RoboDK station: Car_Painting_Cell_v16.rdk

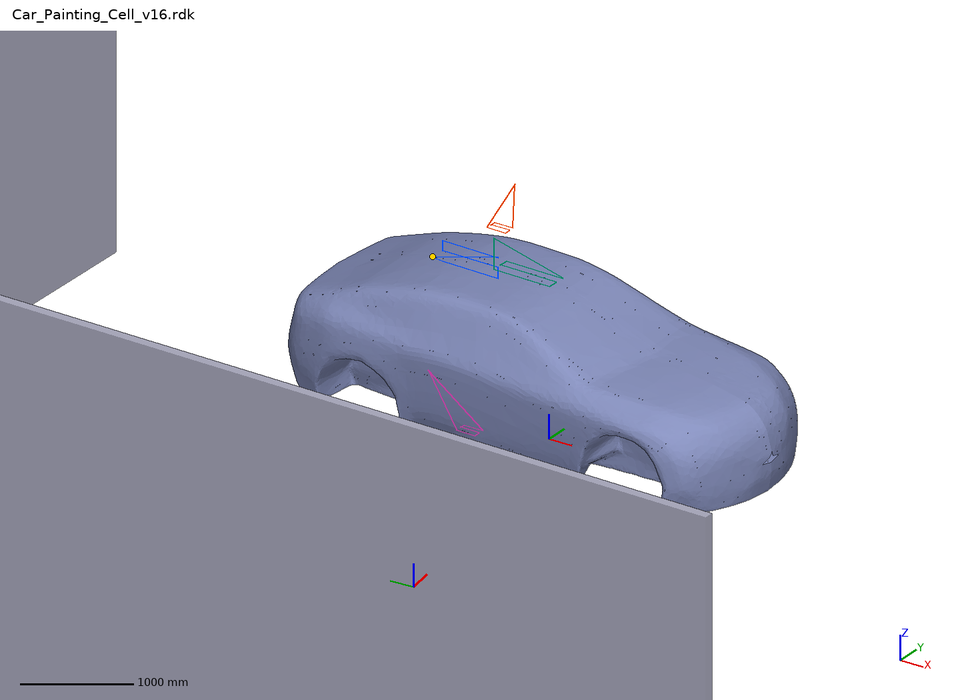
[picture v0: the station drawn from its stored meshes, robots at their saved joint values, targets as dots, program paths as lines]
Station Car_Painting_Cell_v16 (saved by RoboDK 6.1.1). Poses are relative to the parent item; angles as X-Y-Z fixed-axis rotations.
  - frame ABB IRB 6700-235/2.65 Base at (0, 0, 0) mm, rotated rx 1.67 ry -4.75 rz 96.19 deg
    - robot ABB IRB 6700-235/2.65: 6 axes, payload 235 kg, reach 2650 mm, repeatability 0.05 mm, weight 1280 kg
        joint limits [-170, -65, -180, -300, -130, -360] to [170, 85, 70, 300, 130, 360]; home [0, 0, 0, 0, 0, 0]; saved at [22.213, -18.762, 12.242, 0, 96.52, 202.213]
      - tool Generic Paint Sprayer, TCP at (50, 0, 450) mm, rotated rx 0 ry 30 rz 0 deg, size 277.6 x 203.2 x 501.7 mm
  - object Wall_Back at (0, -4050, 2000) mm, size 12000 x 100 x 4000 mm, geometry from Wall_Back.stl
  - object Wall_Side at (-6050, 0, 2000) mm, size 100 x 8000 x 4000 mm, geometry from Wall_Side.stl
  - frame Car_Frame at (-258.38, 2438.18, 404.41) mm
    - object Car_Body at (2438.35, -1259.55, -51.4) mm, rotated rx 0 ry 0 rz 90 deg, size 1981.5 x 4799.5 x 1349.6 mm, geometry from Sedan Car Body.IGS
  - Python program Setup_Cell (listed below)
  - program Paint_Side5 (10 instructions, listed below)
  - program Paint_Trunk2 (10 instructions, listed below)
  - program Paint_Roof2 (10 instructions, listed below)
  - program Paint_Hood2 (10 instructions, listed below)
  - program Main_Program (5 instructions, listed below)
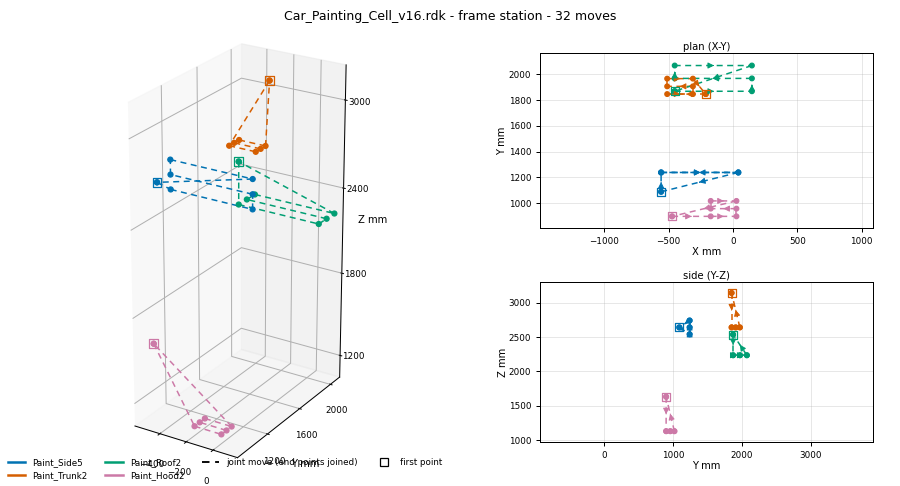
[picture p0: tool path of Car_Painting_Cell_v16.rdk in frame station, 32 of 35 moves have a stored position in this frame; points joined in program order, loops and branches not executed]

--- Python program Setup_Cell ---
# Type help("robodk.robolink") or help("robodk.robomath") for more information
# Press F5 to run the script
# Documentation: https://robodk.com/doc/en/RoboDK-API.html
# Reference:     https://robodk.com/doc/en/PythonAPI/robodk.html
# Note: It is not required to keep a copy of this file, your Python script is saved with your RDK project

# You can also use the new version of the API:
from robodk import robolink    # RoboDK API
from robodk import robomath    # Robot toolbox
RDK = robolink.Robolink()

# Forward and backwards compatible use of the RoboDK API:
# Remove these 2 lines to follow python programming guidelines
from robodk import *      # RoboDK API
from robolink import *    # Robot toolbox
# Link to RoboDK
# RDK = Robolink()

# Notify user:
print('To edit this program:\nright click on the Python program, then, select "Edit Python script"')

# Program example:
item = RDK.Item('base')
if item.Valid():
    print('Item selected: ' + item.Name())
    print('Item posistion: ' + repr(item.Pose()))

print('Items in the station:')
itemlist = RDK.ItemList()
print(itemlist)

# Provoking an exception will display the console output if you run this script from RoboDK
raise Exception('Program not edited.')

--- program Paint_Side5 (robot ABB IRB 6700-235/2.65) ---
  Set Ref.: Car_Frame
  Set Tool: Generic Paint Sprayer
  MoveJ 2 to (-300, -1350, 2235.34) mm, rotated rx -168.9 ry 64.7 rz -87.2 deg; joints [28.216, -32.938, 21.44, 101.638, -42.225, -113.719]
  MoveJ 3 to (-300, -1200, 2135.34) mm, rotated rx -168.9 ry 64.7 rz -87.2 deg; joints [23.122, -28.793, 24.985, 93.784, -36.162, -102.736]
  MoveJ 4 to (300, -1200, 2135.34) mm, rotated rx -168.9 ry 64.7 rz -87.2 deg; joints [-15.84, -33.97, 26.391, 23.272, 7.322, -30.496]
  MoveJ 5 to (300, -1200, 2235.34) mm, rotated rx -168.9 ry 64.7 rz -87.2 deg; joints [-15.495, -31.919, 20.419, 13.499, 10.949, -20.661]
  MoveJ 6 to (-300, -1200, 2235.34) mm, rotated rx -168.9 ry 64.7 rz -87.2 deg; joints [23.087, -26.983, 19.068, 99.337, -36.598, -109.625]
  MoveJ 7 to (-300, -1200, 2335.34) mm, rotated rx -168.9 ry 64.7 rz -87.2 deg; joints [23.052, -24.869, 12.83, 104.706, -37.424, -116.339]
  MoveJ 8 to (300, -1200, 2335.34) mm, rotated rx -168.9 ry 64.7 rz -87.2 deg; joints [-15.156, -29.592, 14.142, 8.67, 14.765, -15.792]
  MoveJ 9 to (-300, -1350, 2235.34) mm, rotated rx -168.9 ry 64.7 rz -87.2 deg; joints [28.216, -32.938, 21.44, 101.638, -42.225, -113.719]

--- program Paint_Trunk2 (robot ABB IRB 6700-235/2.65) ---
  Set Ref.: Car_Frame
  Set Tool: Generic Paint Sprayer
  MoveJ 2 to (47.14, -590.89, 2735.34) mm, rotated rx 176.1 ry 64.7 rz -87.2 deg; joints [-6.92, 10.197, -37.991, 14.59, 28.576, -12.875]
  MoveJ 3 to (-252.86, -590.89, 2235.34) mm, rotated rx 176.1 ry 64.7 rz -87.2 deg; joints [4.168, -2.249, 2.16, -88.78, 4.169, 88.777]
  MoveJ 4 to (-52.86, -590.89, 2235.34) mm, rotated rx 176.1 ry 64.7 rz -87.2 deg; joints [-3.705, -3.302, 2.796, 82.241, 3.739, -82.224]
  MoveJ 5 to (-52.86, -530.89, 2235.34) mm, rotated rx 176.1 ry 64.7 rz -87.2 deg; joints [-3.81, -0.342, 0.158, 87.229, 3.815, -87.223]
  MoveJ 6 to (-252.86, -530.89, 2235.34) mm, rotated rx 176.1 ry 64.7 rz -87.2 deg; joints [3.756, 0.675, -0.495, 87.264, -3.761, -87.258]
  MoveJ 7 to (-252.86, -470.89, 2235.34) mm, rotated rx 176.1 ry 64.7 rz -87.2 deg; joints [3.375, 3.631, -3.327, 84.87, -3.388, -84.861]
  MoveJ 8 to (-52.86, -470.89, 2235.34) mm, rotated rx 176.1 ry 64.7 rz -87.2 deg; joints [-3.908, 2.644, -2.656, 89.824, 3.908, -89.824]
  MoveJ 9 to (47.14, -590.89, 2735.34) mm, rotated rx 176.1 ry 64.7 rz -87.2 deg; joints [-6.92, 10.197, -37.991, 14.59, 28.576, -12.875]

--- program Paint_Roof2 (robot ABB IRB 6700-235/2.65) ---
  Set Ref.: Car_Frame
  Set Tool: Generic Paint Sprayer
  MoveJ 2 to (-194.48, -569.09, 2130.93) mm, rotated rx 176.1 ry 64.7 rz -87.2 deg; joints [12.275, 4.238, -19.199, -40.125, 19.263, 38.507]
  MoveJ 3 to (-194.48, -569.09, 1830.93) mm, rotated rx 176.1 ry 64.7 rz -87.2 deg; joints [12.149, -1.74, 1.882, 89.341, -12.15, -89.326]
  MoveJ 4 to (405.52, -569.09, 1830.93) mm, rotated rx 176.1 ry 64.7 rz -87.2 deg; joints [-11.823, -4.921, 3.782, 84.574, 11.877, -84.456]
  MoveJ 5 to (405.52, -469.09, 1830.93) mm, rotated rx 176.1 ry 64.7 rz -87.2 deg; joints [-11.459, -0.017, -0.535, 87.282, 11.472, -87.227]
  MoveJ 6 to (-194.48, -469.09, 1830.93) mm, rotated rx 176.1 ry 64.7 rz -87.2 deg; joints [10.99, 2.993, -2.518, 87.553, -11, -87.507]
  MoveJ 7 to (-194.48, -369.09, 1830.93) mm, rotated rx 176.1 ry 64.7 rz -87.2 deg; joints [9.964, 7.843, -7.423, 87.611, -9.973, -87.575]
  MoveJ 8 to (405.52, -369.09, 1830.93) mm, rotated rx 176.1 ry 64.7 rz -87.2 deg; joints [-11.141, 4.97, -5.344, 88.1, 11.147, -88.064]
  MoveJ 9 to (-194.48, -569.09, 2130.93) mm, rotated rx 176.1 ry 64.7 rz -87.2 deg; joints [12.275, 4.238, -19.199, -40.125, 19.263, 38.507]

--- program Paint_Hood2 (robot ABB IRB 6700-235/2.65) ---
  Set Ref.: Car_Frame
  Set Tool: Generic Paint Sprayer
  MoveJ 2 to (-214.56, -1541.03, 1228.51) mm, rotated rx -177.97 ry -34.74 rz 95.17 deg; joints [22.213, -18.762, 12.242, 0, 96.52, 202.213]
  MoveJ 3 to (85.44, -1541.03, 728.51) mm, rotated rx -177.97 ry -34.74 rz 95.17 deg; joints [6.355, -29.581, 42.34, 0, 77.241, 186.355]
  MoveJ 4 to (285.44, -1541.03, 728.51) mm, rotated rx -177.97 ry -34.74 rz 95.17 deg; joints [-5.696, -30.968, 42.703, 0, 78.266, 174.304]
  MoveJ 5 to (285.44, -1481.03, 728.51) mm, rotated rx -177.97 ry -34.74 rz 95.17 deg; joints [-5.735, -27.388, 41.004, 0, 76.384, 174.265]
  MoveJ 6 to (85.44, -1481.03, 728.51) mm, rotated rx -177.97 ry -34.74 rz 95.17 deg; joints [5.614, -26.095, 40.626, 0, 75.469, 185.614]
  MoveJ 7 to (85.44, -1421.03, 728.51) mm, rotated rx -177.97 ry -34.74 rz 95.17 deg; joints [4.953, -22.666, 38.771, 0, 73.894, 184.953]
  MoveJ 8 to (285.44, -1421.03, 728.51) mm, rotated rx -177.97 ry -34.74 rz 95.17 deg; joints [-5.769, -23.873, 39.16, 0, 74.713, 174.231]
  MoveJ 9 to (-214.56, -1541.03, 1228.51) mm, rotated rx -177.97 ry -34.74 rz 95.17 deg; joints [22.213, -18.762, 12.242, 0, 96.52, 202.213]

--- program Main_Program (robot ABB IRB 6700-235/2.65) ---
  MoveJ 0 to (0, 0, 0) mm; joints [0, 0, 0, 0, 0, 0]
  Call Paint_Side5
  MoveJ 2 to (0, 0, 0) mm; joints [0, 0, 0, 0, 0, 0]
  Call Paint_Roof2
  MoveJ 4 to (0, 0, 0) mm; joints [0, 0, 0, 0, 0, 0]
